SUBAPPLICATION AX_SoftkeySR_TO_QXA_BG (* 3 Softkeys (SET/RESET/TOGGLE) auf AX_T_FF_SR, Ausgang QXA + Background (am TOGGLE-Key). Generisch. *)
  (* Standard: 61499-2 *)
  (* Version 1.0, 2026-09-09, Franz Höpfinger, Meisterschulen am Ostbahnhof, Ausgelagert aus Uebung_010e2_sub_AX zur Wiederverwendung; u16ObjId_SET/_RESET/_TOGGLE und Output zuvor fest importiert (SoftKey_F1/F2/F3, Output_Q1), jetzt generische Defaults (ID_NULL/Invalid). *)
  PACKAGE MyLib::sys;
  IMPORT isobus::UT::Q::const::IDs::ID_NULL;
  IMPORT logiBUS::io::DQ::logiBUS_DO;
  IMPORT logiBUS::io::DQ::logiBUS_DO_S;
  IMPORT isobus::UT::io::Softkey::SoftKeyActivationCode::SK_RELEASED;
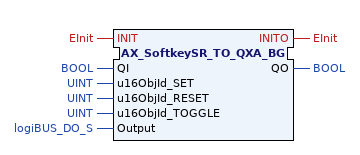
  EVENT_INPUT
    INIT : EInit; (* Initialization Request *)
  END_EVENT
  EVENT_OUTPUT
    INITO : EInit; (* Initialization Confirm *)
  END_EVENT
  VAR_INPUT
    QI : BOOL := TRUE; (* Quality Input - TRUE to enable service *)
    u16ObjId_SET : UINT := ID_NULL; (* Object ID SET SoftKey *)
    u16ObjId_RESET : UINT := ID_NULL; (* Object ID RESET SoftKey *)
    u16ObjId_TOGGLE : UINT := ID_NULL; (* Object ID TOGGLE SoftKey (auch fuer GreenWhiteBackground) *)
    Output : logiBUS::io::DQ::logiBUS_DO_S := logiBUS_DO::Invalid; (* Identify the Output Output_Q1..Q8 *)
  END_VAR
  VAR_OUTPUT
    QO : BOOL; (* Quality Output - TRUE if service executed successfully *)
  END_VAR
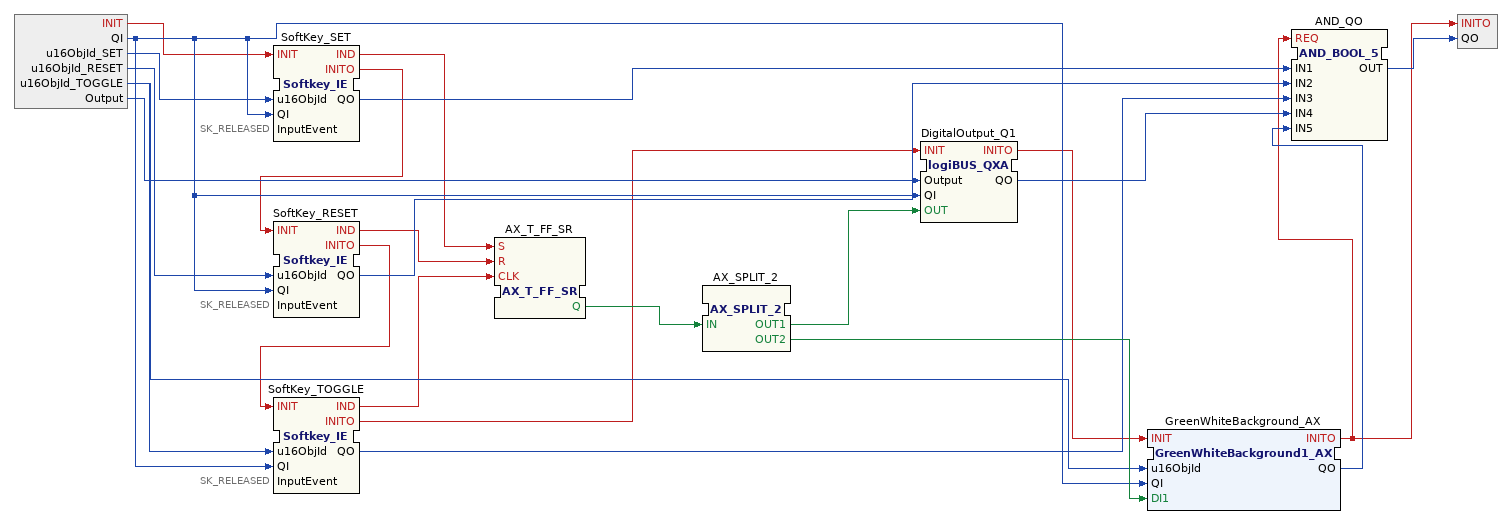
  FBS
    SoftKey_SET : isobus::UT::io::Softkey::Softkey_IE(InputEvent := SK_RELEASED);
    SoftKey_RESET : isobus::UT::io::Softkey::Softkey_IE(InputEvent := SK_RELEASED);
    SoftKey_TOGGLE : isobus::UT::io::Softkey::Softkey_IE(InputEvent := SK_RELEASED);
    AX_T_FF_SR : adapter::events::unidirectional::AX_T_FF_SR;
    AX_SPLIT_2 : adapter::events::unidirectional::AX_SPLIT_2;
    DigitalOutput_Q1 : logiBUS::io::DQ::logiBUS_QXA;
    AND_QO : iec61131::booleanOperators::AND_BOOL_5;
  END_FBS
  SUBAPPS
    GreenWhiteBackground_AX : MyLib::sys::GreenWhiteBackground1_AX;
  END_SUBAPPS
  EVENT_CONNECTIONS
    SoftKey_SET.IND TO AX_T_FF_SR.S;
    SoftKey_RESET.IND TO AX_T_FF_SR.R;
    SoftKey_TOGGLE.IND TO AX_T_FF_SR.CLK;
    INIT TO SoftKey_SET.INIT;
    SoftKey_SET.INITO TO SoftKey_RESET.INIT;
    SoftKey_RESET.INITO TO SoftKey_TOGGLE.INIT;
    SoftKey_TOGGLE.INITO TO DigitalOutput_Q1.INIT;
    DigitalOutput_Q1.INITO TO GreenWhiteBackground_AX.INIT;
    GreenWhiteBackground_AX.INITO TO INITO;
    GreenWhiteBackground_AX.INITO TO AND_QO.REQ;
  END_CONNECTIONS
  DATA_CONNECTIONS
    u16ObjId_SET TO SoftKey_SET.u16ObjId;
    u16ObjId_RESET TO SoftKey_RESET.u16ObjId;
    u16ObjId_TOGGLE TO SoftKey_TOGGLE.u16ObjId;
    u16ObjId_TOGGLE TO GreenWhiteBackground_AX.u16ObjId;
    Output TO DigitalOutput_Q1.Output;
    QI TO SoftKey_SET.QI;
    QI TO SoftKey_RESET.QI;
    QI TO SoftKey_TOGGLE.QI;
    QI TO DigitalOutput_Q1.QI;
    SoftKey_SET.QO TO AND_QO.IN1;
    SoftKey_RESET.QO TO AND_QO.IN2;
    SoftKey_TOGGLE.QO TO AND_QO.IN3;
    DigitalOutput_Q1.QO TO AND_QO.IN4;
    AND_QO.OUT TO QO;
    QI TO GreenWhiteBackground_AX.QI;
    GreenWhiteBackground_AX.QO TO AND_QO.IN5;
  END_CONNECTIONS
  ADAPTER_CONNECTIONS
    AX_T_FF_SR.Q TO AX_SPLIT_2.IN;
    AX_SPLIT_2.OUT1 TO DigitalOutput_Q1.OUT;
    AX_SPLIT_2.OUT2 TO GreenWhiteBackground_AX.DI1;
  END_CONNECTIONS
END_SUBAPPLICATION
